FUNCTION_BLOCK SKILL_Param_INT (* One parameter of a skill: keeps its default, checks a value a client sends with Start against the limits, and holds the value for the run. Technical: Skill parameter (INT): default, range check of a Start argument, latching for one run *)
  (* Standard: 61499-2 *)
  (* Version 0.1, 2026-09-28, Project contributors, AAU Smart Production Lab *)
  PACKAGE modlib;
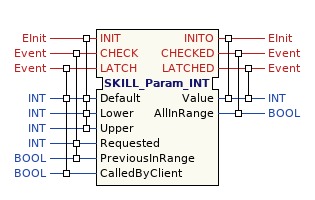
  EVENT_INPUT
    INIT : EInit WITH Default, Lower, Upper; (* Publish the default as the value *)
    CHECK WITH Requested, PreviousInRange; (* Check Requested against Lower..Upper *)
    LATCH WITH CalledByClient, Default; (* Take the value for this run: Requested if CalledByClient, else Default *)
  END_EVENT
  EVENT_OUTPUT
    INITO : EInit WITH Value; (* Initialised: Value is the default *)
    CHECKED WITH AllInRange; (* Checked: AllInRange *)
    LATCHED WITH Value; (* Value holds this run's value *)
  END_EVENT
  VAR_INPUT
    Default : INT; (* The value when the caller gives none; a parent's binding sets it *)
    Lower : INT := -32768; (* The smallest value accepted *)
    Upper : INT := 32767; (* The largest value accepted *)
    Requested : INT; (* The value the caller asks for (an argument of Start) *)
    PreviousInRange : BOOL := TRUE; (* The parameters checked before this one are all in range (TRUE for the first) *)
    CalledByClient : BOOL; (* Started over OPC UA: take Requested, not the default *)
  END_VAR
  VAR_OUTPUT
    Value : INT; (* The value for this run *)
    AllInRange : BOOL; (* This and every parameter before it are in range *)
  END_VAR
  EC_STATES
    INIT : INIT -> INITO;
    CHECK : CHECK -> CHECKED;
    LATCH : LATCH -> LATCHED;
  END_STATES
  ALGORITHM INIT IN ST:
Value := Default;
  END_ALGORITHM
  ALGORITHM CHECK IN ST:
AllInRange := PreviousInRange AND (Requested >= Lower) AND (Requested <= Upper);
  END_ALGORITHM
  ALGORITHM LATCH IN ST:
IF CalledByClient THEN
  Value := Requested;
ELSE
  Value := Default;
END_IF;
  END_ALGORITHM
END_FUNCTION_BLOCK
